(* IEC 61131-3 sources: BODAS-HelloWorld/st/bodas_rc18_12_40/plc_logic/application/03_privatelibrary/datatypes/isobusj1939, 7 files *)

(* ---- enu_isobusj1939_isobusinst-enu_IsobusJ1939_IsobusInst.st ---- *)
(* --- Interface --- *)
{attribute 'qualified_only'}
{attribute 'strict'}
TYPE enu_IsobusJ1939_IsobusInst : (
		IsobusJ1939_IsobusInst1_E := 1, (* FOR CAN1 *)
		IsobusJ1939_IsobusInst2_E := 2, (* for CAN2 *)
		IsobusJ1939_IsobusInst3_E := 3, (* for CAN3 *)
		IsobusJ1939_IsobusInstMax_E     (* last enum for automatic array resizing *)
	);
END_TYPE

(* ---- enu_isobusj1939_rxinst1box-enu_IsobusJ1939_RxInst1Box.st ---- *)
(* --- Interface --- *)
{attribute 'qualified_only'}
{attribute 'strict'}
TYPE enu_IsobusJ1939_RxInst1Box : (
		IsobusJ1939_RxInst1BoxDm1_E := 3,
		IsobusJ1939_RxInst1BoxMax_E (* last enum for automatic array resizing *)
	);
END_TYPE

(* ---- enu_isobusj1939_rxinst2box-enu_IsobusJ1939_RxInst2Box.st ---- *)
(* --- Interface --- *)
{attribute 'qualified_only'}
{attribute 'strict'}
TYPE enu_IsobusJ1939_RxInst2Box : (
		IsobusJ1939_RxInst2BoxDm1_E := 3,
		IsobusJ1939_RxInst2BoxMax_E (* last enum for automatic array resizing *)
	);
END_TYPE

(* ---- enu_isobusj1939_rxinst3box-enu_IsobusJ1939_RxInst3Box.st ---- *)
(* --- Interface --- *)
{attribute 'qualified_only'}
{attribute 'strict'}
TYPE enu_IsobusJ1939_RxInst3Box : (
		IsobusJ1939_RxInst3BoxDm1_E := 3,
		IsobusJ1939_RxInst3BoxMax_E (* last enum for automatic array resizing *)
	);
END_TYPE

(* ---- enu_isobusj1939_txinst1box-enu_IsobusJ1939_TxInst1Box.st ---- *)
(* --- Interface --- *)
{attribute 'qualified_only'}
{attribute 'strict'}
TYPE enu_IsobusJ1939_TxInst1Box : (
		IsobusJ1939_TxInst1BoxDm1_E := 3,
		IsobusJ1939_TxInst1BoxDm2_E,
		IsobusJ1939_TxInst1BoxDummy1Tx_E,
		IsobusJ1939_TxInst1BoxMax_E (* last enum for automatic array resizing *)
	);
END_TYPE

(* ---- enu_isobusj1939_txinst2box-enu_IsobusJ1939_TxInst2Box.st ---- *)
(* --- Interface --- *)
{attribute 'qualified_only'}
{attribute 'strict'}
TYPE enu_IsobusJ1939_TxInst2Box : (
		IsobusJ1939_TxInst2BoxDm1_E := 3,
		IsobusJ1939_TxInst2BoxMax_E (* last enum for automatic array resizing *)
	);
END_TYPE

(* ---- enu_isobusj1939_txinst3box-enu_IsobusJ1939_TxInst3Box.st ---- *)
(* --- Interface --- *)
{attribute 'qualified_only'}
{attribute 'strict'}
TYPE enu_IsobusJ1939_TxInst3Box : (
		IsobusJ1939_TxInst3BoxDm1_E := 3,
		IsobusJ1939_TxInst3BoxMax_E (* last enum for automatic array resizing *)
	);
END_TYPE
